FUNCTION_BLOCK Magazine1 (* Composite Function Block Type *)
  (* Standard: 61499-2 *)
  (* Version 0.0, 7/2/2026, template *)
  PACKAGE Main;
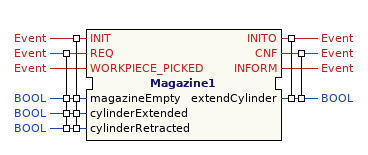
  EVENT_INPUT
    INIT WITH magazineEmpty, cylinderExtended, cylinderRetracted; (* Initialization Request *)
    REQ WITH magazineEmpty, cylinderExtended, cylinderRetracted; (* Normal Execution Request *)
    WORKPIECE_PICKED;
  END_EVENT
  EVENT_OUTPUT
    INITO WITH extendCylinder; (* Initialization Confirm *)
    CNF WITH extendCylinder; (* Execution Confirmation *)
    INFORM;
  END_EVENT
  VAR_INPUT
    magazineEmpty : BOOL; (* Input event qualifier *)
    cylinderExtended : BOOL;
    cylinderRetracted : BOOL;
  END_VAR
  VAR_OUTPUT
    extendCylinder : BOOL; (* Output event qualifier *)
  END_VAR
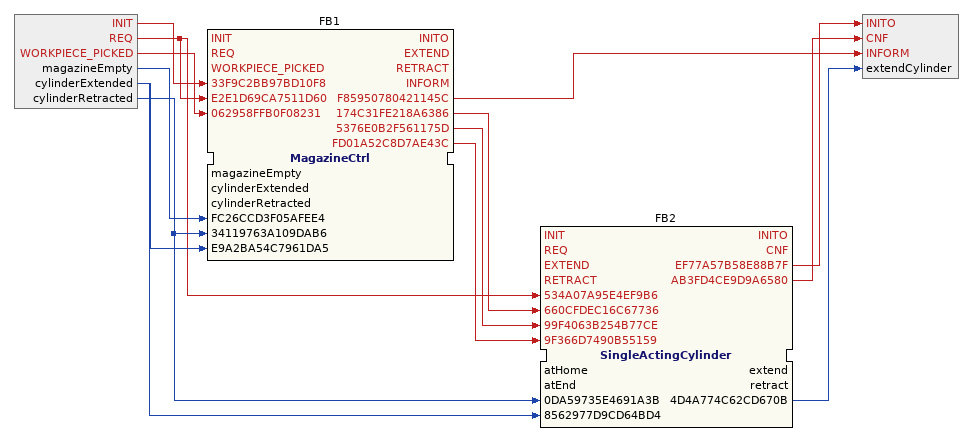
  FBS
    FB1 : MagazineCtrl;
    FB2 : SingleActingCylinder;
  END_FBS
  EVENT_CONNECTIONS
    FB2.EF77A57B58E88B7F TO INITO;
    FB2.AB3FD4CE9D9A6580 TO CNF;
    FB1.F85950780421145C TO INFORM;
    INIT TO FB1.33F9C2BB97BD10F8;
    REQ TO FB1.E2E1D69CA7511D60;
    REQ TO FB2.534A07A95E4EF9B6;
    WORKPIECE_PICKED TO FB1.062958FFB0F08231;
    FB1.174C31FE218A6386 TO FB2.660CFDEC16C67736;
    FB1.5376E0B2F561175D TO FB2.99F4063B254B77CE;
    FB1.FD01A52C8D7AE43C TO FB2.9F366D7490B55159;
  END_CONNECTIONS
  DATA_CONNECTIONS
    FB2.4D4A774C62CD670B TO extendCylinder;
    magazineEmpty TO FB1.FC26CCD3F05AFEE4;
    cylinderRetracted TO FB1.34119763A109DAB6;
    cylinderRetracted TO FB2.0DA59735E4691A3B;
    cylinderExtended TO FB1.E9A2BA54C7961DA5;
    cylinderExtended TO FB2.8562977D9CD64BD4;
  END_CONNECTIONS
END_FUNCTION_BLOCK
